(* IEC 61131-3 sources: llm-plc-st-eval/data/processed_definitivo/gemini-3.1-pro-preview/A4/zero_shot, 3 files *)

(* ---- ejec_1.st ---- *)
FUNCTION_BLOCK FB_Rampa
VAR_INPUT
    SPvel : REAL;       (* Consigna de velocidad *)
    paroRapido : BOOL;  (* Comando de paro rápido *)
    ciclo : TIME;       (* Tiempo de ciclo de ejecución del bloque *)
END_VAR

VAR_OUTPUT
    CVvel : REAL;       (* Velocidad actual de salida *)
END_VAR

VAR
    ciclo_s : REAL;     (* Tiempo de ciclo convertido a segundos *)
    target : REAL;      (* Valor objetivo temporal *)
    tasa : REAL;        (* Tasa de cambio activa (%/s) *)
    delta_max : REAL;   (* Cambio máximo permitido en el ciclo actual *)
    diferencia : REAL;  (* Diferencia entre el objetivo y la salida actual *)
END_VAR

(* Convertir el tiempo de ciclo (TIME) a segundos (REAL) *)
(* Se asume que TIME_TO_UDINT devuelve el tiempo en milisegundos, estándar en IEC 61131-3 *)
ciclo_s := UDINT_TO_REAL(TIME_TO_UDINT(ciclo)) / 1000.0;

(* Determinar el objetivo y la tasa de cambio según el estado *)
IF paroRapido THEN
    target := 0.0;
    tasa := 40.0;       (* Pendiente de paro rápido *)
ELSE
    target := SPvel;
    IF target > CVvel THEN
        tasa := 10.0;   (* Pendiente de subida *)
    ELSIF target < CVvel THEN
        tasa := 20.0;   (* Pendiente de bajada *)
    ELSE
        tasa := 0.0;    (* Sin cambio *)
    END_IF;
END_IF;

(* Calcular el incremento máximo y la diferencia *)
delta_max := tasa * ciclo_s;
diferencia := target - CVvel;

(* Actualizar la salida evitando el sobrepaso *)
IF ABS(diferencia) <= delta_max THEN
    CVvel := target;                (* Alcanza el objetivo sin sobrepasarlo *)
ELSIF diferencia > 0.0 THEN
    CVvel := CVvel + delta_max;     (* Incrementa hacia el objetivo *)
ELSE
    CVvel := CVvel - delta_max;     (* Decrementa hacia el objetivo *)
END_IF;

END_FUNCTION_BLOCK

(* ---- ejec_2.st ---- *)
FUNCTION_BLOCK FB_Rampa
VAR_INPUT
    SPvel : REAL;       (* Consigna de velocidad objetivo *)
    paroRapido : BOOL;  (* Comando para detención rápida *)
    ciclo : TIME;       (* Período de ejecución del bloque *)
END_VAR

VAR_OUTPUT
    CVvel : REAL;       (* Velocidad de salida con rampa aplicada *)
END_VAR

VAR
    dt : REAL;          (* Tiempo de ciclo convertido a segundos *)
    objetivo : REAL;    (* Valor al que debe tender la salida *)
    deltaMax : REAL;    (* Cambio máximo permitido en el ciclo actual *)
    diferencia : REAL;  (* Diferencia entre el objetivo y la salida actual *)
END_VAR

(* 1. Convertir el tiempo de ciclo (TIME) a segundos (REAL) *)
dt := TIME_TO_REAL(ciclo) / 1000.0;

(* 2. Determinar el valor objetivo y el incremento/decremento máximo (deltaMax) *)
IF paroRapido THEN
    objetivo := 0.0;
    deltaMax := 40.0 * dt; (* Pendiente de paro rápido: 40.0 %/s *)
ELSE
    objetivo := SPvel;
    IF objetivo > CVvel THEN
        deltaMax := 10.0 * dt; (* Pendiente de subida normal: 10.0 %/s *)
    ELSE
        deltaMax := 20.0 * dt; (* Pendiente de bajada normal: 20.0 %/s *)
    END_IF;
END_IF;

(* 3. Calcular la diferencia entre el objetivo y el valor actual *)
diferencia := objetivo - CVvel;

(* 4. Aplicar la rampa asegurando que no haya sobrepaso *)
IF diferencia > 0.0 THEN
    (* Se requiere subir la velocidad *)
    IF diferencia > deltaMax THEN
        CVvel := CVvel + deltaMax;
    ELSE
        CVvel := objetivo; (* Evita el sobrepaso *)
    END_IF;
ELSIF diferencia < 0.0 THEN
    (* Se requiere bajar la velocidad *)
    IF -diferencia > deltaMax THEN
        CVvel := CVvel - deltaMax;
    ELSE
        CVvel := objetivo; (* Evita el sobrepaso *)
    END_IF;
END_IF;

END_FUNCTION_BLOCK

(* ---- ejec_3.st ---- *)
FUNCTION_BLOCK FB_Rampa
VAR_INPUT
    SPvel : REAL;       (* Consigna de velocidad objetivo *)
    paroRapido : BOOL;  (* Comando de paro rápido *)
    ciclo : TIME;       (* Período de ejecución del bloque *)
END_VAR
VAR_OUTPUT
    CVvel : REAL;       (* Consigna de velocidad actual (salida con rampa) *)
END_VAR
VAR
    ciclo_s : REAL;     (* Tiempo de ciclo convertido a segundos *)
    target : REAL;      (* Objetivo de velocidad a alcanzar *)
    stepUp : REAL;      (* Paso máximo de incremento por ciclo *)
    stepDown : REAL;    (* Paso máximo de decremento por ciclo *)
END_VAR

(* Convertir el tiempo de ciclo a segundos (asumiendo que TIME internamente está en milisegundos) *)
ciclo_s := DINT_TO_REAL(TIME_TO_DINT(ciclo)) / 1000.0;

(* Configurar el objetivo y las pendientes según el estado de paro rápido *)
IF paroRapido THEN
    target := 0.0;
    (* En paro rápido, la pendiente es 40.0 pts/s tanto si desciende desde positivo como si asciende desde negativo *)
    stepUp := 40.0 * ciclo_s;
    stepDown := 40.0 * ciclo_s;
ELSE
    target := SPvel;
    stepUp := 10.0 * ciclo_s;   (* Pendiente de subida: 10.0 pts/s *)
    stepDown := 20.0 * ciclo_s; (* Pendiente de bajada: 20.0 pts/s *)
END_IF;

(* Aplicar la rampa hacia el objetivo asegurando que no haya sobrepaso *)
IF CVvel < target THEN
    CVvel := CVvel + stepUp;
    IF CVvel > target THEN
        CVvel := target; (* Evitar sobrepaso al subir *)
    END_IF;
ELSIF CVvel > target THEN
    CVvel := CVvel - stepDown;
    IF CVvel < target THEN
        CVvel := target; (* Evitar sobrepaso al bajar *)
    END_IF;
END_IF;

END_FUNCTION_BLOCK
